(*
SPDX-FileCopyrightText: © 2026 Oleksandr Tiutyk <trofimich@gmail.com>
SPDX-License-Identifier: MIT
License: https://opensource.org/license/mit
*)

(*!
<summary>Holds long text and a distinct marker for native capacity and encoding tests.</summary>
*)
TYPE JSON_TEST_LARGE_VALUE :
STRUCT
	//! <summary>Uses the framework JSON text capacity in bytes, excluding the terminator.</summary>
	Text : STRING(TOF_Core.Parameters.JSON_DOCUMENT_CHAR_SIZE);
	//! <summary>Independent field that distinguishes the structure from its first member.</summary>
	Marker : DINT;
END_STRUCT
END_TYPE

(* stored: Version 1.1.0.1
   DUT JSON_TEST_LARGE_VALUE: Id {c0f7b9f1-a78e-49c9-a8a8-8ea2e8f6dda4} *)
